// Transfer function RPM <-> PWM duty cycle.
// RpmLow corresponds to 0 %, RpmHigh to 100 %. The result is limited to 0..100 %.
// RpmHigh < RpmLow is allowed and inverts the characteristic.
FUNCTION_BLOCK RpmToDutyCycle IMPLEMENTS I_TransformLRealValue
VAR
	_RpmLow	 : LREAL := 0.0;
	_RpmHigh : LREAL := 1000.0;
END_VAR
VAR CONSTANT
	DUTY_CYCLE_MIN : LREAL := 10.0;
	DUTY_CYCLE_MAX : LREAL := 90.0;
END_VAR

PROPERTY RpmHigh : LREAL // RPM at 100 % duty cycle
GET // PUBLIC
RpmHigh := _RpmHigh;
END_GET
SET // PUBLIC
_RpmHigh := RpmHigh;
END_SET
END_PROPERTY

PROPERTY RpmLow : LREAL // RPM at 0 % duty cycle
GET // PUBLIC
RpmLow := _RpmLow;
END_GET
SET // PUBLIC
_RpmLow := RpmLow;
END_SET
END_PROPERTY

// Reverse = FALSE: RPM -> duty cycle [%]
// Reverse = TRUE : duty cycle [%] -> RPM
// Returns 0 if RpmLow = RpmHigh (invalid range).
METHOD Transform : LREAL
VAR_INPUT
	Value	: LREAL;
    Reverse : BOOL := FALSE;
END_VAR
VAR
	Span : LREAL;
END_VAR
Span := _RpmHigh - _RpmLow;
IF Span = 0.0 THEN
	Transform := 0.0;
	RETURN;
END_IF

IF NOT Reverse THEN
	// RPM -> duty cycle [%]: RpmLow..RpmHigh maps to DUTY_CYCLE_MIN..DUTY_CYCLE_MAX
	IF Value <= _RpmLow THEN
		Transform := DUTY_CYCLE_MIN;
	ELSIF Value >= _RpmHigh THEN
		Transform := DUTY_CYCLE_MAX;
	ELSE
		Transform := DUTY_CYCLE_MIN + (Value - _RpmLow) / Span * (DUTY_CYCLE_MAX - DUTY_CYCLE_MIN);
	END_IF
ELSE
	// Duty cycle [%] -> RPM: DUTY_CYCLE_MIN..DUTY_CYCLE_MAX maps to RpmLow..RpmHigh
	IF Value <= DUTY_CYCLE_MIN THEN
		Transform := _RpmLow;
	ELSIF Value >= DUTY_CYCLE_MAX THEN
		Transform := _RpmHigh;
	ELSE
		Transform := _RpmLow + (Value - DUTY_CYCLE_MIN) / (DUTY_CYCLE_MAX - DUTY_CYCLE_MIN) * Span;
	END_IF
END_IF
END_METHOD

END_FUNCTION_BLOCK

(* stored: Version 1.1.0.1
   POU RpmToDutyCycle: Id {6df2fede-0591-457a-93f9-83fe478b07b8}, SpecialFunc None
   Property RpmHigh: Id {69f01143-a1a9-4f8b-a21f-4d8ab8421ef9}
   Get Get: Id {a8ee8911-02fb-40bd-920d-a61a073baa17}
   Set Set: Id {a2950738-a557-46f8-b8bb-842ea46192f1}
   Property RpmLow: Id {213e2254-3340-4321-a14c-3f0458586ff5}
   Get Get: Id {f28aad5b-6f30-4dd9-b706-99a3d46e938e}
   Set Set: Id {34b2de77-0ebe-46d5-a933-f3059496660a}
   Method Transform: Id {007c82bf-5092-4835-93c6-a62f349e2dfc} *)
